(* ============================================================
   GVL_SML_CONST - LIBRARY constants (invariants)
   SML

   Only constants owned by the library (machine-independent).
   The application configuration (number of axes) lives in GVL_App.MAX_AXIS.
   Qualified reference: GVL_SML_CONST.PROGRESS_SPAN, ...
   ============================================================ *)

{attribute 'qualified_only'}
VAR_GLOBAL CONSTANT
    PROGRESS_SPAN : DINT := 100;   // progress band width in the combined state
                                   // (E_AXIS_STATE values are multiples of this)

    // -- MAPPING: fixed size (bytes) of the bus blocks for the UNIONs --
    // Must be >= SIZEOF of the corresponding struct (checked at runtime
    // by FB_Mapping_In/Out via Check). Fixed for a stable process image
    // on the fieldbus.
    MAP_SIZE_CTRL  : UDINT := 64;    // >= SIZEOF(ST_AXIS_CTRL)
    MAP_SIZE_DATA  : UDINT := 64;    // >= SIZEOF(ST_MOVE_DATA)
    MAP_SIZE_STATE : UDINT := 256;   // >= SIZEOF(ST_AXIS_STATE) (holds 2x STRING(80))
    MAP_SIZE_INFO  : UDINT := 128;   // >= SIZEOF(ST_AXIS_INFO) (with Status + TouchProbe)
END_VAR

(* stored: Version 1.1.0.1
   GVL GVL_SML_CONST: Id {12bf8a46-3177-54ca-8f1a-432f6a0d29c7} *)
